// TIA Portal V19 export
TYPE "UDT_TachoDT_Q"
   STRUCT
      TSV_102 : Bool;   // Soplo de vapor directo al cuerpo
      XSV_112B : Bool;   // Meladura cruda: vÃ¡lvula de rama al cabezal comÃºn
      XSV_112A : Bool;   // Meladura clara: vÃ¡lvula de rama al cabezal comÃºn
      XSV_105 : Bool;   // AlimentaciÃ³n de semilla
      PSV_103 : Bool;   // RompevacÃ­o / admisiÃ³n de aire
      LSV_109 : Bool;   // Descarga de masa cocida al recibidor
      XSV_104 : Bool;   // InyecciÃ³n de colada
      XSV_108 : Bool;   // Transferencia Tacho 3 -> Tacho 2
      M_101 : Bool;   // Motor agitador
      XSV_113 : Bool;   // Drenaje (reserva/futuro)
      M_102 : Bool;   // Bomba de vacÃ­o Consignas analÃ³gicas de vÃ¡lvulas: RAW 0..27648 = 0..100 %
      LCV_212_RAW : Int;   // AlimentaciÃ³n comÃºn de meladuras
      DCV_211_RAW : Int;   // Vapor a calandria
      XCV_107_RAW : Int;   // Agua caliente al cuerpo
      PCV_210_RAW : Int;   // Agua de enfriamiento al condensador
   END_STRUCT;
END_TYPE
